// TIA Portal V19 export
// export: Created 2026-10-15T09:44:24.0910042Z, ExportSetting WithDefaults, DisplayName Totally Integrated Automation Portal, DisplayVersion V19, DisplayName TIA Portal Openness, DisplayVersion V19, DisplayName TIA Portal Version Control Interface, DisplayVersion V19, DisplayName STEP 7 Professional, DisplayVersion V19, DisplayName STEP 7 Safety, DisplayVersion V19, DisplayName WinCC Basic/Comfort/Advanced, DisplayVersion V19, DisplayName WinCC Unified, DisplayVersion V19
FUNCTION "ROLL_PB13" : Void   // FC21, SCL
{ S7_Optimized_Access := 'TRUE' }
VERSION : 0.1
// stored: AutoNumber true, IsIECCheckEnabled false, SetENOAutomatically false, UDAEnableTagReadback false
   VAR_TEMP
      r : Bool;
      a1 : Word;
      a2 : Word;
      activeDataBlock : Int;
      comparisonResults : Array[0..0] of Bool;
   END_VAR
BEGIN

   #r := FALSE;
   #a1 := W#16#0000;
   #a2 := W#16#0000;
   #activeDataBlock := 0;
   // PB13, STEP 5 network 1
   #r := ((NOT "ROLL_State".M[58, 6]) AND ("ROLL_IO".Input[11, 1] OR "ROLL_IO".Input[11, 2] OR "ROLL_IO".Input[11, 3] OR "ROLL_IO".Input[11, 4] OR "ROLL_IO".Input[119, 6] OR "ROLL_IO".Input[119, 7] OR "ROLL_IO".Input[120, 0]) AND "ROLL_IO".Input[11, 6]);
   IF #r THEN
       "ROLL_State".M[58, 7] := TRUE;
   END_IF;
   #r := (((NOT "ROLL_IO".Input[11, 6]) AND ("ROLL_IO".Input[11, 1] OR "ROLL_IO".Input[11, 2] OR "ROLL_IO".Input[11, 3] OR "ROLL_IO".Input[11, 4] OR "ROLL_IO".Input[119, 6] OR "ROLL_IO".Input[119, 7] OR "ROLL_IO".Input[120, 0]) AND "ROLL_IO".Output[23, 0] AND "ROLL_State".M[58, 6]) OR "ROLL_IO".Input[11, 0]);
   IF #r THEN
       "ROLL_State".M[58, 7] := FALSE;
   END_IF;
   // PB13, STEP 5 network 2
   #r := "ROLL_IO".Input[11, 6];
   "ROLL_State".M[58, 6] := #r;
   // PB13, STEP 5 network 3
   #r := (((((NOT "ROLL_IO".Input[11, 0]) OR "ROLL_State".M[80, 7]) AND "ROLL_IO".Input[11, 6]) OR "ROLL_State".M[58, 7]) AND "ROLL_IO".Input[14, 0]);
   "ROLL_State".M[60, 0] := #r;
   // PB13, STEP 5 network 4
   #a2 := #a1;
   #a1 := W#16#2030;
   #r := ((NOT "ROLL_IO".Input[13, 3]) AND "ROLL_IO".Output[24, 0]);
   "ROLL_TimerOp"(Number := 110,
                  Operation := 0,
                  Signal := #r,
                  Preset := #a1);
   // PB13, STEP 5 network 5
   #r := (((NOT "ROLL_State".M[111, 1]) AND (NOT "ROLL_State".M[111, 2]) AND (NOT "ROLL_State".M[111, 5]) AND "ROLL_IO".Input[0, 2] AND "ROLL_State".M[111, 0]) OR ((NOT "ROLL_State".M[61, 5]) AND "ROLL_IO".Input[0, 1] AND "ROLL_State".M[23, 2]) OR ("ROLL_IO".Input[12, 1] AND "ROLL_State".M[111, 5]));
   "ROLL_State".M[60, 1] := #r;
   // PB13, STEP 5 network 6
   #r := (((NOT "ROLL_IO".Input[12, 1]) AND "ROLL_State".M[111, 5]) OR ((NOT "ROLL_State".M[111, 0]) AND (NOT "ROLL_State".M[111, 2]) AND (NOT "ROLL_State".M[111, 5]) AND "ROLL_IO".Input[0, 2] AND "ROLL_State".M[111, 1]) OR ("ROLL_IO".Input[0, 1] AND "ROLL_State".M[23, 3]));
   "ROLL_State".M[60, 3] := #r;
   // PB13, STEP 5 network 7
   #r := (((NOT "ROLL_State".M[111, 0]) AND (NOT "ROLL_State".M[111, 1]) AND (NOT "ROLL_State".M[111, 5]) AND "ROLL_IO".Input[0, 2] AND "ROLL_State".M[111, 2]) OR ((NOT "ROLL_State".M[61, 5]) AND "ROLL_IO".Input[0, 1] AND "ROLL_State".M[0, 3]));
   "ROLL_State".M[60, 2] := #r;
   // PB13, STEP 5 network 8
   #a2 := #a1;
   #a1 := W#16#0005;
   #r := (NOT "ROLL_State".S5Timers[114].Q);
   "ROLL_TimerOp"(Number := 113,
                  Operation := 0,
                  Signal := #r,
                  Preset := #a1);
   #a2 := #a1;
   #a1 := W#16#0005;
   #r := "ROLL_State".S5Timers[113].Q;
   "ROLL_TimerOp"(Number := 114,
                  Operation := 1,
                  Signal := #r,
                  Preset := #a1);
   // PB13, STEP 5 network 9
   #activeDataBlock := 15;
   // PB13, STEP 5 network 10
   #a2 := #a1;
   #a1 := "ROLL_GetDW"(DbNumber := #activeDataBlock, Index := 116);
   #r := ((NOT "ROLL_State".S5Timers[117].Q) AND "ROLL_State".M[62, 4]);
   "ROLL_TimerOp"(Number := 116,
                  Operation := 0,
                  Signal := #r,
                  Preset := #a1);
   #a2 := #a1;
   #a1 := "ROLL_GetDW"(DbNumber := #activeDataBlock, Index := 117);
   #r := "ROLL_State".S5Timers[116].Q;
   "ROLL_TimerOp"(Number := 117,
                  Operation := 1,
                  Signal := #r,
                  Preset := #a1);
   // PB13, STEP 5 network 11
   #activeDataBlock := 19;
   // PB13, STEP 5 network 12
   #r := ("ROLL_IO".Output[24, 2] AND "ROLL_State".M[60, 4] AND "ROLL_State".S5Timers[114].Q);
   "ROLL_CounterOp"(Number := 1,
                    Operation := 3,
                    Signal := #r,
                    Preset := #a1);
   #a2 := #a1;
   #a1 := "ROLL_GetDW"(DbNumber := #activeDataBlock, Index := 1);
   #r := ((((NOT "ROLL_IO".Input[13, 3]) AND (NOT ("ROLL_State".S5Counters[1].Value <> 0)) AND (NOT ("ROLL_State".S5Counters[2].Value <> 0))) OR "ROLL_IO".Input[13, 3] OR "ROLL_State".M[60, 5]) AND "ROLL_State".S5Timers[114].Q);
   "ROLL_CounterOp"(Number := 1,
                    Operation := 0,
                    Signal := #r,
                    Preset := #a1);
   // PB13, STEP 5 network 13
   #r := ("ROLL_IO".Output[24, 0] AND "ROLL_State".M[60, 5] AND "ROLL_State".S5Timers[114].Q);
   "ROLL_CounterOp"(Number := 2,
                    Operation := 3,
                    Signal := #r,
                    Preset := #a1);
   #a2 := #a1;
   #a1 := "ROLL_GetDW"(DbNumber := #activeDataBlock, Index := 2);
   #r := (("ROLL_IO".Input[13, 3] OR "ROLL_State".M[60, 4]) AND "ROLL_State".S5Timers[114].Q);
   "ROLL_CounterOp"(Number := 2,
                    Operation := 0,
                    Signal := #r,
                    Preset := #a1);
   // PB13, STEP 5 network 14
   #r := ((NOT "ROLL_IO".Input[13, 3]) AND "ROLL_IO".Output[24, 2] AND "ROLL_State".M[60, 6]);
   IF #r THEN
       "ROLL_State".M[60, 4] := TRUE;
   END_IF;
   #r := "ROLL_IO".Input[13, 3];
   IF #r THEN
       "ROLL_State".M[60, 4] := FALSE;
   END_IF;
   // PB13, STEP 5 network 15
   #r := ((NOT "ROLL_IO".Input[13, 3]) AND "ROLL_IO".Output[24, 0] AND "ROLL_State".M[60, 6]);
   IF #r THEN
       "ROLL_State".M[60, 5] := TRUE;
   END_IF;
   #r := "ROLL_IO".Input[13, 3];
   IF #r THEN
       "ROLL_State".M[60, 5] := FALSE;
   END_IF;
   // PB13, STEP 5 network 16
   #r := "ROLL_IO".Input[13, 3];
   IF #r THEN
       "ROLL_State".M[60, 6] := TRUE;
   END_IF;
   #r := ("ROLL_State".M[60, 4] OR "ROLL_State".M[60, 5]);
   IF #r THEN
       "ROLL_State".M[60, 6] := FALSE;
   END_IF;
   // PB13, STEP 5 network 17
   #r := ((NOT ("ROLL_State".S5Counters[2].Value <> 0)) AND "ROLL_State".M[62, 6]);
   IF #r THEN
       "ROLL_State".M[60, 7] := TRUE;
   END_IF;
   #r := (NOT "ROLL_State".M[62, 6]);
   IF #r THEN
       "ROLL_State".M[60, 7] := FALSE;
   END_IF;
   // PB13, STEP 5 network 18
   #r := ((NOT "ROLL_IO".Input[13, 3]) AND (NOT ("ROLL_State".S5Counters[1].Value <> 0)) AND "ROLL_State".M[61, 1]);
   IF #r THEN
       "ROLL_State".M[61, 0] := TRUE;
   END_IF;
   #r := (NOT "ROLL_State".M[62, 6]);
   IF #r THEN
       "ROLL_State".M[61, 0] := FALSE;
   END_IF;
   // PB13, STEP 5 network 19
   #r := ("ROLL_State".S5Counters[1].Value <> 0);
   "ROLL_State".M[61, 1] := #r;
   // PB13, STEP 5 network 20
   #r := (("ROLL_State".M[60, 7] OR "ROLL_State".M[62, 6]) AND "ROLL_State".M[61, 0]);
   "ROLL_State".M[61, 2] := #r;
   // PB13, STEP 5 network 21
   #r := ((NOT "ROLL_State".M[61, 6]) AND "ROLL_State".M[60, 1] AND "ROLL_State".M[61, 7]);
   IF #r THEN
       "ROLL_State".M[61, 3] := TRUE;
   END_IF;
   #r := (NOT "ROLL_State".M[61, 7]);
   IF #r THEN
       "ROLL_State".M[61, 3] := FALSE;
   END_IF;
   // PB13, STEP 5 network 22
   #r := ((NOT "ROLL_State".M[61, 6]) AND "ROLL_State".M[60, 2] AND "ROLL_State".M[61, 7]);
   IF #r THEN
       "ROLL_State".M[61, 4] := TRUE;
   END_IF;
   #r := (NOT "ROLL_State".M[61, 7]);
   IF #r THEN
       "ROLL_State".M[61, 4] := FALSE;
   END_IF;
   // PB13, STEP 5 network 23
   #r := ((NOT "ROLL_State".M[61, 6]) AND "ROLL_State".M[60, 3] AND "ROLL_State".M[61, 7]);
   IF #r THEN
       "ROLL_State".M[61, 5] := TRUE;
   END_IF;
   #r := (NOT "ROLL_State".M[61, 7]);
   IF #r THEN
       "ROLL_State".M[61, 5] := FALSE;
   END_IF;
   // PB13, STEP 5 network 24
   #r := "ROLL_State".M[61, 7];
   "ROLL_State".M[61, 6] := #r;
   // PB13, STEP 5 network 25
   #r := (((NOT "ROLL_State".M[111, 5]) AND "ROLL_State".M[37, 3]) OR ((((NOT "ROLL_IO".Input[12, 1]) AND ("ROLL_State".M[41, 0] OR "ROLL_State".M[42, 4] OR "ROLL_State".M[44, 0])) OR (("ROLL_State".M[40, 5] OR "ROLL_State".M[42, 1] OR "ROLL_State".M[43, 5]) AND "ROLL_IO".Input[12, 1])) AND "ROLL_State".M[111, 5]));
   IF #r THEN
       "ROLL_State".M[61, 7] := TRUE;
   END_IF;
   #r := (((NOT "ROLL_IO".Input[12, 5]) AND "ROLL_IO".Input[11, 0] AND "ROLL_State".M[190, 5] AND "ROLL_State".M[20, 1]) OR (("ROLL_State".M[42, 0] OR "ROLL_State".M[43, 4] OR "ROLL_State".M[58, 5]) AND "ROLL_State".M[111, 5]) OR "ROLL_State".M[53, 6]);
   IF #r THEN
       "ROLL_State".M[61, 7] := FALSE;
   END_IF;
   // PB13, STEP 5 network 26
   #r := ((NOT "ROLL_IO".Input[11, 0]) AND (((NOT "ROLL_IO".Input[12, 1]) AND "ROLL_IO".Output[23, 5]) OR ("ROLL_IO".Output[23, 4] AND "ROLL_IO".Input[12, 1])) AND ("ROLL_State".M[61, 3] OR "ROLL_State".M[61, 4] OR "ROLL_State".M[61, 5]));
   IF #r THEN
       "ROLL_State".M[62, 0] := TRUE;
   END_IF;
   #r := ((("ROLL_State".M[41, 3] OR "ROLL_State".M[42, 7] OR "ROLL_State".M[44, 3] OR "ROLL_State".M[46, 0] OR "ROLL_State".M[47, 3] OR "ROLL_State".M[48, 7] OR "ROLL_State".M[50, 3] OR "ROLL_State".M[51, 5]) AND "ROLL_IO".Input[13, 3] AND "ROLL_State".S5Timers[114].Q) OR (NOT "ROLL_State".M[31, 5]) OR (NOT "ROLL_State".M[61, 7]));
   IF #r THEN
       "ROLL_State".M[62, 0] := FALSE;
   END_IF;
   // PB13, STEP 5 network 27
   #r := (((NOT "ROLL_IO".Input[11, 0]) AND ((("ROLL_IO".Input[11, 1] OR "ROLL_IO".Input[11, 2] OR "ROLL_IO".Input[11, 3] OR "ROLL_IO".Input[11, 4] OR "ROLL_IO".Input[119, 6] OR "ROLL_IO".Input[119, 7] OR "ROLL_IO".Input[120, 0]) AND ("ROLL_State".M[80, 6] OR "ROLL_State".M[80, 7])) OR ("ROLL_State".M[60, 0] AND "ROLL_State".M[80, 7]))) OR ("ROLL_IO".Input[11, 0] AND "ROLL_IO".Input[11, 6] AND "ROLL_State".M[80, 7]));
   "ROLL_State".M[62, 1] := #r;
   // PB13, STEP 5 network 28
   #r := (("ROLL_State".M[0, 3] AND "ROLL_State".M[45, 6]) OR "ROLL_State".M[41, 1] OR "ROLL_State".M[42, 5] OR "ROLL_State".M[44, 1] OR "ROLL_State".M[47, 1] OR "ROLL_State".M[48, 5] OR "ROLL_State".M[50, 1]);
   "ROLL_State".M[63, 5] := #r;
   // PB13, STEP 5 network 29
   #r := (((((NOT "ROLL_State".M[60, 1]) AND (NOT "ROLL_State".M[60, 2]) AND (NOT "ROLL_State".M[60, 3]) AND (NOT "ROLL_State".M[63, 1]) AND "ROLL_State".M[74, 0]) OR ((NOT "ROLL_State".M[60, 1]) AND (NOT "ROLL_State".M[60, 2]) AND "ROLL_State".M[60, 3])) AND ("ROLL_State".M[20, 1] OR "ROLL_State".M[20, 2] OR "ROLL_State".M[23, 3]) AND "ROLL_IO".Input[0, 1]) OR ((((NOT "ROLL_State".M[61, 3]) AND (NOT "ROLL_State".M[61, 4]) AND (NOT "ROLL_State".M[61, 5]) AND "ROLL_State".M[62, 6]) OR ((NOT "ROLL_State".M[61, 3]) AND (NOT "ROLL_State".M[61, 4]) AND "ROLL_State".M[61, 5])) AND "ROLL_IO".Input[0, 2]));
   "ROLL_State".M[62, 2] := #r;
   // PB13, STEP 5 network 30
   #r := (((NOT "ROLL_State".M[60, 2]) AND (NOT "ROLL_State".M[60, 3]) AND ("ROLL_State".M[20, 1] OR "ROLL_State".M[23, 2]) AND "ROLL_IO".Input[0, 1] AND "ROLL_State".M[60, 1]) OR ((NOT "ROLL_State".M[61, 4]) AND (NOT "ROLL_State".M[61, 5]) AND (NOT "ROLL_State".M[63, 5]) AND "ROLL_IO".Input[0, 2] AND "ROLL_State".M[61, 3]));
   "ROLL_State".M[62, 3] := #r;
   // PB13, STEP 5 network 31
   #r := (((NOT "ROLL_State".M[60, 1]) AND (NOT "ROLL_State".M[60, 3]) AND ("ROLL_State".M[0, 3] OR "ROLL_State".M[20, 1]) AND "ROLL_IO".Input[0, 1] AND "ROLL_State".M[60, 2]) OR ((((NOT "ROLL_State".M[61, 3]) AND (NOT "ROLL_State".M[61, 5]) AND "ROLL_State".M[61, 4]) OR ("ROLL_State".M[61, 3] AND "ROLL_State".M[63, 5])) AND "ROLL_IO".Input[0, 2]));
   "ROLL_State".M[62, 4] := #r;
   // PB13, STEP 5 network 32
   #r := ((((NOT "ROLL_State".M[190, 5]) AND ("ROLL_State".M[0, 3] OR "ROLL_State".M[23, 2] OR "ROLL_State".M[23, 3]) AND ("ROLL_State".M[60, 1] OR "ROLL_State".M[60, 2] OR "ROLL_State".M[60, 3]) AND "ROLL_IO".Input[0, 1] AND "ROLL_State".M[190, 6] AND "ROLL_State".M[62, 1]) OR ("ROLL_IO".Input[0, 2] AND "ROLL_State".M[31, 5] AND "ROLL_State".M[62, 0])) AND ("ROLL_State".M[62, 5] OR "ROLL_State".S5Timers[114].Q) AND "ROLL_State".M[60, 0]);
   "ROLL_State".M[62, 5] := #r;
   // PB13, STEP 5 network 33
   #r := ((NOT "ROLL_State".M[63, 1]) AND (((NOT "ROLL_State".M[62, 0]) AND "ROLL_IO".Input[0, 2] AND "ROLL_State".M[31, 5]) OR ((((NOT "ROLL_State".M[190, 6]) AND ("ROLL_State".M[0, 3] OR "ROLL_State".M[20, 2] OR "ROLL_State".M[23, 2] OR "ROLL_State".M[23, 3]) AND "ROLL_State".M[190, 5]) OR "ROLL_State".M[74, 0]) AND "ROLL_IO".Input[0, 1] AND "ROLL_State".M[62, 1])) AND ("ROLL_State".M[62, 6] OR "ROLL_State".S5Timers[114].Q) AND "ROLL_State".M[60, 0]);
   "ROLL_State".M[62, 6] := #r;
   // PB13, STEP 5 network 34
   #r := ((((NOT "ROLL_State".M[61, 2]) AND (NOT "ROLL_State".M[63, 1]) AND "ROLL_State".M[62, 6]) OR "ROLL_State".M[62, 5]) AND (((NOT "ROLL_State".M[62, 2]) AND (NOT "ROLL_State".M[62, 4]) AND (NOT "ROLL_State".M[62, 6]) AND "ROLL_State".M[62, 3]) OR ((NOT "ROLL_State".M[62, 6]) AND ("ROLL_IO".Input[13, 3] OR "ROLL_State".S5Timers[117].Q) AND "ROLL_State".M[62, 4]) OR (((NOT "ROLL_State".M[62, 4]) OR "ROLL_State".M[62, 6]) AND ("ROLL_State".S5Counters[1].Value <> 0))) AND ("ROLL_State".M[62, 2] OR "ROLL_State".M[62, 3] OR "ROLL_State".M[62, 4]));
   "ROLL_State".M[62, 7] := #r;
   // PB13, STEP 5 network 35
   #r := ((NOT "ROLL_IO".Output[24, 0]) AND (NOT "ROLL_State".M[5, 1]) AND (NOT "ROLL_State".M[63, 4]) AND ((NOT "ROLL_State".S5Timers[115].Q) OR "ROLL_IO".Output[24, 2]) AND "ROLL_IO".Input[13, 5] AND "ROLL_State".M[29, 0] AND "ROLL_State".M[60, 0] AND "ROLL_State".M[62, 7]);
   "ROLL_IO".Output[24, 2] := #r;
   // PB13, STEP 5 network 36
   #r := ((((NOT "ROLL_State".M[62, 2]) AND (NOT "ROLL_State".M[62, 6])) OR ("ROLL_State".S5Counters[2].Value <> 0)) AND (((NOT "ROLL_State".M[63, 1]) AND "ROLL_State".M[62, 6]) OR "ROLL_State".M[62, 5]) AND ((NOT "ROLL_State".M[62, 4]) OR (NOT "ROLL_State".M[62, 5])));
   "ROLL_State".M[63, 0] := #r;
   // PB13, STEP 5 network 37
   #r := ((NOT "ROLL_IO".Output[24, 2]) AND (NOT "ROLL_State".M[5, 1]) AND (NOT "ROLL_State".M[63, 4]) AND ((NOT "ROLL_State".S5Timers[115].Q) OR "ROLL_IO".Output[24, 0]) AND "ROLL_IO".Input[13, 5] AND "ROLL_State".M[29, 0] AND "ROLL_State".M[60, 0] AND "ROLL_State".M[63, 0]);
   "ROLL_IO".Output[24, 0] := #r;
   // PB13, STEP 5 network 38
   #r := ((NOT "ROLL_IO".Output[24, 5]) AND "ROLL_IO".Output[24, 0] AND "ROLL_IO".Input[13, 3]);
   "ROLL_IO".Output[24, 1] := #r;
   // PB13, STEP 5 network 39
   #r := ("ROLL_IO".Output[24, 0] OR "ROLL_IO".Output[24, 2] OR "ROLL_State".M[63, 6]);
   "ROLL_State".M[240, 0] := #r;
   // PB13, STEP 5 network 40
   #r := ((NOT "ROLL_IO".Input[12, 5]) AND (("ROLL_State".M[190, 5] AND "ROLL_State".M[23, 0]) OR "ROLL_State".M[52, 2]) AND "ROLL_IO".Input[11, 0] AND "ROLL_IO".Input[11, 6]);
   IF #r THEN
       "ROLL_State".M[63, 6] := TRUE;
   END_IF;
   #r := (("ROLL_IO".Input[12, 1] OR "ROLL_IO".Input[12, 5]) AND "ROLL_IO".Input[11, 0] AND "ROLL_IO".Input[11, 6] AND "ROLL_IO".Input[12, 7]);
   IF #r THEN
       "ROLL_State".M[63, 6] := FALSE;
   END_IF;
   // PB13, STEP 5 network 41
   #r := ((((NOT "ROLL_State".M[63, 7]) AND "ROLL_IO".Output[24, 0] AND "ROLL_State".S5Timers[111].Q) OR ("ROLL_IO".Input[11, 0] AND "ROLL_State".M[80, 6]) OR (NOT "ROLL_State".S5Timers[11].Q)) AND "ROLL_IO".Input[13, 3]);
   IF #r THEN
       "ROLL_State".M[63, 1] := TRUE;
   END_IF;
   #r := (((NOT "ROLL_IO".Input[13, 3]) AND "ROLL_IO".Input[3, 0] AND "ROLL_State".S5Timers[11].Q) OR "ROLL_IO".Output[24, 2]);
   IF #r THEN
       "ROLL_State".M[63, 1] := FALSE;
   END_IF;
   // PB13, STEP 5 network 42
   #a2 := #a1;
   #a1 := W#16#1030;
   #r := ("ROLL_IO".Output[24, 0] AND "ROLL_IO".Input[13, 3] AND "ROLL_State".M[29, 0] AND "ROLL_State".M[61, 2]);
   "ROLL_TimerOp"(Number := 111,
                  Operation := 0,
                  Signal := #r,
                  Preset := #a1);
   // PB13, STEP 5 network 43
   #r := (((NOT "ROLL_IO".Input[13, 3]) AND "ROLL_IO".Input[0, 1] AND "ROLL_State".M[0, 3] AND "ROLL_State".M[190, 6]) OR ((((NOT "ROLL_State".M[61, 2]) AND "ROLL_State".M[62, 6]) OR "ROLL_State".M[62, 5]) AND ("ROLL_State".M[62, 2] OR "ROLL_State".M[62, 3] OR "ROLL_State".M[62, 4])) OR ("ROLL_IO".Input[13, 3] AND "ROLL_State".M[63, 7]));
   "ROLL_State".M[63, 7] := #r;
   "ROLL_IO".Output[24, 5] := #r;
   // PB13, STEP 5 network 44
   #r := ("ROLL_IO".Output[24, 0] OR "ROLL_IO".Output[24, 2]);
   "ROLL_IO".Output[24, 4] := #r;
   // PB13, STEP 5 network 45
   #r := ("ROLL_State".M[41, 1] OR "ROLL_State".M[42, 5] OR "ROLL_State".M[44, 1] OR "ROLL_State".M[45, 6] OR "ROLL_State".M[47, 1] OR "ROLL_State".M[48, 5] OR "ROLL_State".M[50, 1]);
   "ROLL_State".M[240, 0] := #r;
   // PB13, STEP 5 network 46
   #r := "ROLL_State".M[111, 1];
   "ROLL_State".M[240, 1] := #r;
   // PB13, STEP 5 network 47
   "ROLL_FB69"();
   // PB13, STEP 5 network 48
   #a2 := #a1;
   #a1 := "ROLL_GetM"(FirstByte := 240, Width := 16);
   #r := ("ROLL_IO".Output[24, 0] OR "ROLL_IO".Output[24, 2]);
   "ROLL_TimerOp"(Number := 115,
                  Operation := 1,
                  Signal := #r,
                  Preset := #a1);
   // PB13, STEP 5 network 49
   #r := ((("ROLL_IO".Output[24, 0] AND "ROLL_State".M[60, 5]) OR ("ROLL_IO".Output[24, 2] AND "ROLL_State".M[60, 4])) AND "ROLL_State".S5Timers[114].Q);
   "ROLL_CounterOp"(Number := 3,
                    Operation := 3,
                    Signal := #r,
                    Preset := #a1);
   #r := ((((NOT "ROLL_State".M[60, 4]) AND (NOT "ROLL_State".M[60, 5]) AND ("ROLL_IO".Output[24, 0] OR "ROLL_IO".Output[24, 2])) OR ("ROLL_IO".Output[24, 0] AND "ROLL_State".M[60, 4]) OR ("ROLL_IO".Output[24, 2] AND "ROLL_State".M[60, 5])) AND "ROLL_State".S5Timers[114].Q);
   "ROLL_CounterOp"(Number := 3,
                    Operation := 2,
                    Signal := #r,
                    Preset := #a1);
   #a2 := #a1;
   #a1 := W#16#0500;
   #r := (("ROLL_IO".Input[13, 3] AND "ROLL_State".S5Timers[114].Q) OR ("ROLL_State".M[3, 1] AND "ROLL_State".M[63, 2]));
   "ROLL_CounterOp"(Number := 3,
                    Operation := 0,
                    Signal := #r,
                    Preset := #a1);
   // PB13, STEP 5 network 50
   #a2 := #a1;
   #a1 := INT_TO_WORD("ROLL_State".S5Counters[3].Value);
   #a2 := #a1;
   #a1 := W#16#0208;
   #comparisonResults[0] := (WORD_TO_INT(#a2) > WORD_TO_INT(#a1));
   #r := #comparisonResults[0];
   "ROLL_State".M[63, 2] := #r;
   // PB13, STEP 5 network 51
   #a2 := #a1;
   #a1 := W#16#1060;
   #r := ((("ROLL_IO".Output[24, 0] AND "ROLL_State".M[63, 7]) OR "ROLL_IO".Output[24, 2]) AND "ROLL_IO".Input[13, 3]);
   "ROLL_TimerOp"(Number := 112,
                  Operation := 0,
                  Signal := #r,
                  Preset := #a1);
   // PB13, STEP 5 network 52
   #r := ((NOT ("ROLL_State".S5Counters[2].Value <> 0)) AND "ROLL_State".M[61, 2] AND "ROLL_State".M[62, 6] AND ("ROLL_State".S5Counters[1].Value <> 0));
   "ROLL_State".M[63, 3] := #r;
   // PB13, STEP 5 network 53
   #r := (((NOT "ROLL_IO".Input[0, 4]) AND "ROLL_IO".Input[0, 2] AND "ROLL_State".M[63, 4]) OR "ROLL_State".M[11, 0] OR "ROLL_State".M[11, 1] OR "ROLL_State".M[11, 2] OR "ROLL_State".M[11, 3]);
   "ROLL_State".M[63, 4] := #r;
   // PB13, STEP 5 network 54
   RETURN;
END_FUNCTION
